(* IEC 61131-3 sources: plc-iiot-stack/tools/tests/fixtures/sample/src/Interfaces/I_Resettable, 1 file *)

(* ---- Reset.method.decl.st ---- *)
// Сброс; TRUE — отказ сброшен
METHOD Reset : BOOL
VAR_INPUT
    xForce : BOOL;  // сброс без проверки условий
END_VAR
